Staubli VAL3: click_logSave.pgx

program click_logSave()
  local num l_nResult
  local string l_sDate
begin
  //  l_sDate=getDate("%m_%d %H_%M_%S")
  //  call rs:saveLog("./LOG_"+l_sDate,l_nResult)
  call rs:saveLog(""+l_sDate,l_nResult)
  if l_nResult!=0
    popUpMsg("保存失败:"+toString("",l_nResult))
    return
  endIf
  popUpMsg("保存成功")
end
